// Base of the CFC test suites. TcUnit's TEST and TEST_FINISHED_NAMED are functions without a return
// type, which a CFC box cannot call (the editor insists on a return pin), so the diagrams call these
// two methods instead. Everything else comes from TcUnit.FB_TestSuite.
FUNCTION_BLOCK ABSTRACT T_SafeCfcTestSuite EXTENDS TcUnit.FB_TestSuite

// Marks the start of a test (TcUnit.TEST). Call it first in every test method, every cycle.
METHOD PROTECTED StartTest
VAR_INPUT
    TestName : T_MaxString;
END_VAR
TcUnit.TEST(TestName);
END_METHOD

// Marks a test as finished (TcUnit.TEST_FINISHED_NAMED).
METHOD PROTECTED FinishTest
VAR_INPUT
    TestName : T_MaxString;
END_VAR
TcUnit.TEST_FINISHED_NAMED(TestName);
END_METHOD

END_FUNCTION_BLOCK

(* stored: Version 1.1.0.1, ProductVersion 3.1.4026.22
   POU T_SafeCfcTestSuite: Id {5b8db23e-b89f-53f5-a9dd-2055a694f476}, SpecialFunc None
   Method StartTest: Id {a7b7a387-18ba-56fd-ad9d-c291f19aaaad}
   Method FinishTest: Id {063209f1-29d3-5445-b235-6819f9af0ff8} *)
